// TIA Portal V21 export
// export: Created 2026-11-21T11:47:44.3091465Z, ExportSetting WithDefaults, DisplayName Totally Integrated Automation Portal, DisplayVersion V21, DisplayName STEP 7 Professional, DisplayVersion V21, DisplayName STEP 7 Safety, DisplayVersion V21, DisplayName Tech WebApplication, DisplayVersion V21, DisplayName WinCC Basic/Comfort/Advanced, DisplayVersion V21, DisplayName WinCC Unified, DisplayVersion V21
FUNCTION_BLOCK "LadBoxes"   // FB11, LAD
TITLE = Boxes
{ S7_Optimized_Access := 'TRUE' }
VERSION : 0.1
// Boxes in ladder: move, compare, add, timers, a counter and calls.
// stored: AutoNumber true, IsIECCheckEnabled false, IsRetainMemResEnabled false, MemoryReserve 100, SetENOAutomatically false, UDAEnableTagReadback false
   VAR_INPUT
      level : Int;
      count : Bool;
      reset : Bool;
   END_VAR
   VAR_OUTPUT
      high : Bool;
      clamped : Int;
      done : Bool;
      pulse : Bool;
   END_VAR
   VAR
      delay : TON_TIME;
   END_VAR
   VAR RETAIN
      "counter" : CTU_INT;
   END_VAR
   VAR
      pulser : "Pulse";
      copy : Int;
      sum : Int;
   END_VAR
BEGIN

REGION Network 1: Move
   // Copies the level.
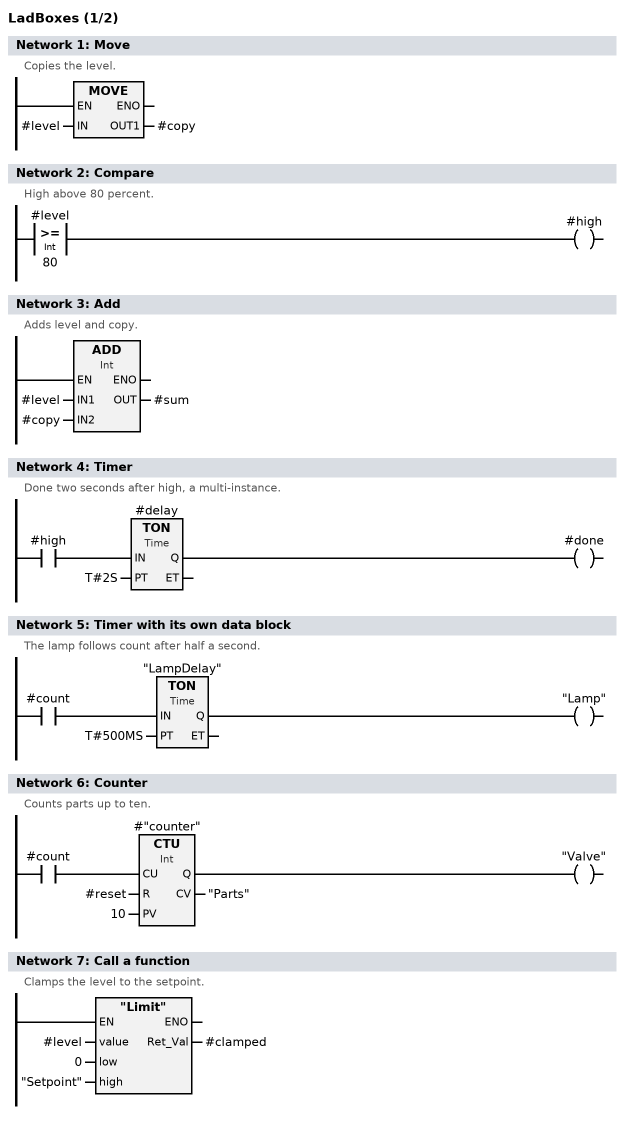
   RUNG wire#powerrail
      { S7_GenerateENO := "TRUE" } Move(in := #level, out1 => #copy)
   END_RUNG
   // the same network as SCL:
   #copy := #level;
END_REGION

REGION Network 2: Compare
   // High above 80 percent.
   RUNG wire#powerrail
      { S7_Templates := "SrcType := Int" } GE_Contact(in1 := #level, in2 := 80)
      Coil( #high )
   END_RUNG
   // the same network as SCL:
   #high := #level >= 80;
END_REGION

REGION Network 3: Add
   // Adds level and copy.
   RUNG wire#powerrail
      { S7_Templates := "SrcType := Int"; S7_GenerateENO := "TRUE" } Add(in1 := #level, in2 := #copy, out => #sum)
   END_RUNG
   // the same network as SCL:
   #sum := #level + #copy;
END_REGION

REGION Network 4: Timer
   // Done two seconds after high, a multi-instance.
   RUNG wire#powerrail
      Contact( #high )
      { S7_Templates := "time_type := Time" } #delay.TON(pt := T#2S, et =>)
      Coil( #done )
   END_RUNG
   // the same network as SCL:
   #delay(IN := #high, PT := T#2S);   // TON
   #done := #delay.Q;
END_REGION

REGION Network 5: Timer with its own data block
   // The lamp follows count after half a second.
   RUNG wire#powerrail
      Contact( #count )
      { S7_Templates := "time_type := Time" } "LampDelay".TON(pt := T#500MS, et =>)
      Coil( "Lamp" )
   END_RUNG
   // the same network as SCL:
   "LampDelay".TON(IN := #count, PT := T#500MS);
   "Lamp" := "LampDelay".Q;
END_REGION

REGION Network 6: Counter
   // Counts parts up to ten.
   RUNG wire#powerrail
      Contact( #count )
      { S7_Templates := "value_type := Int" } #"counter".CTU(r := #reset, pv := 10, cv => "Parts")
      Coil( "Valve" )
   END_RUNG
   // the same network as SCL:
   #"counter"(CU := #count, R := #reset, PV := 10, CV => "Parts");   // CTU
   "Valve" := #"counter".Q;
END_REGION

REGION Network 7: Call a function
   // Clamps the level to the setpoint.
   RUNG wire#powerrail
      "Limit"(value := #level, low := 0, high := "Setpoint", Ret_Val => #clamped)
   END_RUNG
   // the same network as SCL:
   #clamped := "Limit"(value := #level, low := 0, high := "Setpoint");
END_REGION

REGION Network 8: Call a function block
   // A pulse on each count, a multi-instance.
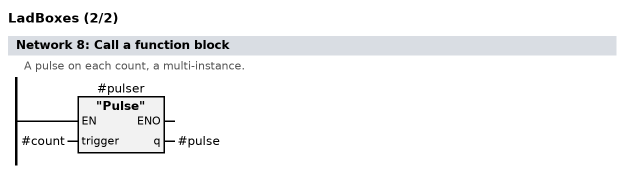
   RUNG wire#powerrail
      #pulser(trigger := #count, q => #pulse)
   END_RUNG
   // the same network as SCL:
   #pulser(trigger := #count, q => #pulse);   // "Pulse"
END_REGION
END_FUNCTION_BLOCK
